(* IEC 61131-3 sources: plc-process-lib/tools/demo/src/POUs/PRG_Demo, 2 files *)

(* ---- PRG_Demo.decl.st ---- *)
// Назначение: программа демонстрационного прогона (задача MainTask, 10 мс): общий отсчёт
//             времени от системного источника библиотеки и три независимых сценария на ФБ
//             plc-process-lib 1.0.0.0 — контур уровня (A), классификация NE 43 (B), тревога
//             ISA-18.2 (C). Устройства берут время сами (itfTime не задан — системное время), то
//             есть прогон идёт в реальном времени. Когда все сценарии завершены — xAllDone.
// Автор:      kr0nsch
// Версия:     0.1.0
// Документ:   docs/media/data/demo-run.json; tools/demo/README.md
PROGRAM PRG_Demo
VAR
    fbClock  : PL.FB_SystemTime;   // системное время библиотеки (монотонное LTIME)
    xStarted : BOOL;               // первый цикл выполнен
    ltStart  : LTIME;              // время старта сценариев
    ltPrev   : LTIME;              // время прошлого цикла
    ltNow    : LTIME;              // время этого цикла
    lrT_s    : LREAL;              // время от старта, с
    lrDt_s   : LREAL;              // шаг цикла, с
    fbLoop   : FB_DemoLevelLoop;   // A: контур уровня
    fbNe43   : FB_DemoNe43;        // B: NE 43
    fbAlarm  : FB_DemoAlarm;       // C: тревога ISA-18.2
END_VAR

(* ---- PRG_Demo.impl.st ---- *)
ltNow := fbClock.Now();
IF NOT xStarted THEN
    xStarted := TRUE;
    ltStart := ltNow;
    ltPrev := ltNow;
END_IF
lrT_s := PL.F_LTimeToSec(ltIn := ltNow - ltStart);
lrDt_s := PL.F_LTimeToSec(ltIn := ltNow - ltPrev);
ltPrev := ltNow;

fbLoop(lrT_s := lrT_s, lrDt_s := lrDt_s);
fbNe43(lrT_s := lrT_s);
fbAlarm(lrT_s := lrT_s);
GVL_DemoLog.xAllDone := fbLoop.xDone AND fbNe43.xDone AND fbAlarm.xDone;
